(* IEC 61131-3 sources: 2026_Projet_YGO_ExcavatriceDragage/CODE/ENCODERS, 5 files *)

(* ---- ST_EncoderCalib.st ---- *)
(* ═══════════════════════════════════════════════════════════════
   🧲 ST_EncoderCalib — Calibration/référence codeur (1 par treuil, RETAIN)
   ───────────────────────────────────────────────────────────────
   📄 Doc métier : DOC/AF_Partie10_Fonction_Encoder_Homing_v1.6.md §9
   🎛️ Une instance RETAIN par treuil (M1_EncoderCalib / M2_EncoderCalib).
   ⚠️ Ce lot (acquisition + mise à l'échelle) : `HomingRefRaw` reste
      modifiable MANUELLEMENT (RETAIN, valeur de test) tant que
      `FB_Encoder_Homing` (qui l'écrit normalement, §5) n'est pas codé —
      même principe que le stub GVL du lot Winch.
   ═══════════════════════════════════════════════════════════════ *)

TYPE ST_EncoderCalib :
STRUCT
    HomingRefRaw                  : UDINT;   // Valeur brute figée au dernier homing réussi
    LastKnownRawPos                : UDINT;   // Dernier point brut valide connu (§3.7, continu)
    RestartCoherenceTolerancePts    : UDINT := 1000;  // Tolérance redémarrage (~12% PointsPerRev 8192)
    Homed                          : BOOL;    // TRUE dès qu'un référencement a réussi
    HomingSuspect                  : BOOL;    // TRUE si incohérence détectée au redémarrage (§3.7)
END_STRUCT
END_TYPE

(* ---- FB_Encoder_Abs.st ---- *)
(* ═══════════════════════════════════════════════════════════════
   🧲 FB_Encoder_Abs — Acquisition codeur absolu (accès bus, 1 responsabilité)
   ───────────────────────────────────────────────────────────────
   📄 Doc métier : DOC/AF_Partie10_Fonction_Encoder_Homing_v1.6.md §3/§6
   ⚠️ RÉÉCRITURE COMPLÈTE (remplace la version legacy du projet, dossier
      CODEUR) : l'ancienne version utilisait `HomingTrigger` (recalage
      instantané par simple offset) + un mode `Teach` auto-calibré —
      **incompatibles** avec le design Partie10 (preset SDO avec
      accusé, formule `CableM_PerRev` fixe). Retirés : `HomingTrigger`,
      `WaterLevelOffset`, `TeachActive/StartRaw/EndRaw/RealDistance`.
   🧩 1 FB = 1 responsabilité : accès bus EtherCAT + séquence d'écriture
      preset. N'orchestre PAS le homing lui-même (ça sera le rôle de
      `FB_Encoder_Homing`, pas codé ce lot) — `PresetRequest`/`PresetValue`
      sont pilotés en dur (`FALSE`/`0`) dans `PRG_MAIN` pour l'instant.
   🧊 Principe « geler sur doute » (§6) : `RawPos`/`AngleRaw`/`TurnCount`
      ne sont PAS mis à jour si `EncoderAvailable = FALSE` — ils
      conservent leur dernière valeur plausible.
   ✅ SÉQUENCE PRESET (§5) — CONFIRMÉ TERRAIN 2026-07-02 : `PresetTriggerCmd := 2`
      (valeur de commande, pas un masque de bits) déclenche le
      référencement du codeur à `PresetValueOut`. `CodeSeqTriggerCmd`
      (canal réel `COD1_CodeSeqTrigCmd`) reste `0`, rôle **non identifié**
      (même par l'utilisateur/terrain) — ne jamais lui donner une valeur
      arbitraire tant que sa fonction n'est pas confirmée.
   🔴 PERTE DE FONCTION SIGNALÉE : l'ancienne version composait
      `FB_Encoder_Safety` en interne (survitesse via `In_SpdValue`).
      Ce n'est PAS repris ici (Partie10 ne le demande pas, hors
      périmètre du document) — `FB_Encoder_Safety` (overspeed) devient
      orphelin tant qu'un lot dédié ne décide pas de son sort (fusion
      avec le "saut incohérent" Partie10 §3.5, ou reprise telle quelle).
   🔧 CORRECTIF (2026-07-03, retour terrain) : `InvertDirection` **retiré**.
      Confirmé terrain : l'objet CoE `6000h` (bit0 : 4→5) inverse le sens
      de comptage **côté codeur** (F58x8 Kübler), configuré en **Startup
      Parameter** CODESYS (init automate) — pas un paramètre PLC. L'ancien
      calcul logiciel (`16#FFFFFFFF - RawPosIn`) était de toute façon
      **buggé** : il inversait sur toute la plage `UDINT` (32 bits) au
      lieu de la plage réelle du codeur (25 bits, `PointsPerRev ×
      MultiTurnRevsMax`), produisant des positions incohérentes après
      homing. Voir Partie10 §3bis.
   ═══════════════════════════════════════════════════════════════ *)

// === DECLARATION (à coller dans la partie déclaration du POU FB_Encoder_Abs) ===

FUNCTION_BLOCK PUBLIC FB_Encoder_Abs
VAR_INPUT
    Enable              : BOOL;        // Standard
    Reset               : BOOL;        // Acquittement défaut (front)
    EmergencyStopOk     : BOOL;        // Standard
    Mode                : E_Mode;      // Standard (contexte, pas encore exploité ce lot)
    RawPosIn            : UDINT;       // Brut EtherCAT (ex. COD1_PosValue, %ID)
    AlarmsIn            : UINT;        // Brut EtherCAT (ex. COD1_Alarms)
    WarningsIn          : UINT;        // Brut EtherCAT (ex. COD1_Warnings) — informatif seulement
    SlaveOperational    : BOOL;        // FB_DiagEthercat — esclave EtherCAT opérationnel
    PointsPerRev        : UDINT := 8192;  // Résolution codeur confirmée (Partie10 §3.3)
    PresetRequest       : BOOL;        // Front — piloté par FB_Encoder_Homing (stub FALSE ce lot)
    PresetValue         : UDINT;       // Cible brute — piloté par FB_Encoder_Homing (stub 0 ce lot)
    PresetTimeout       : TIME := T#2s;
    PresetTolerancePts  : UDINT := 10; // Tolérance relecture post-preset
END_VAR
VAR_OUTPUT
    Ready               : BOOL;
    Busy                : BOOL;
    Done                : BOOL;
    Error               : BOOL;
    ErrorId             : WORD;        // bit0: "Défaut communication codeur" - alarme/bus codeur ; bit1: "Erreur référencement (timeout)" - preset refusé/timeout
    State               : E_State;
    StateAtError        : E_State;
    RawPos              : UDINT;       // Position brute — GELÉE si EncoderAvailable=FALSE
    EncoderAvailable    : BOOL;
    AngleRaw            : UINT;        // Informatif maintenance : RawPos MOD PointsPerRev
    TurnCount           : UDINT;       // Informatif maintenance : RawPos / PointsPerRev
    PresetAck           : BOOL;        // Pulse 1 cycle — écriture confirmée
    PresetNak           : BOOL;        // Pulse 1 cycle — écriture refusée/timeout
    PresetTriggerCmd    : WORD;        // → à câbler sur COD_PresettTrigCmd (RxPDO)
    CodeSeqTriggerCmd   : WORD;        // → à câbler sur COD_CodeSeqTrigCmd (RxPDO)
    PresetValueOut      : UDINT;       // → à câbler sur COD_PresetValue (RxPDO)
END_VAR
VAR
    ResetEdge           : R_TRIG;
    ErrorEdge           : R_TRIG;
    PresetReqEdge       : R_TRIG;
    PresetTimer         : TON;
    PresetSeqStep       : INT;         // 0=IDLE, 1=pulse CodeSeq, 2=pulse Trig, 3=attente confirmation
    RawDiff             : DINT;
    PresetTimerVisual   : TON;         // Timer pour laisser le temps de voir l'impulsion (1.5s)
END_VAR

// === IMPLEMENTATION (à coller dans le corps ST du POU FB_Encoder_Abs) ===

// 🛑 1. GATE
IF NOT Enable THEN
    EncoderAvailable := FALSE;
    State := E_State.DISABLED;
    Ready := FALSE; Busy := FALSE; Done := FALSE;
    PresetTriggerCmd := 16#0000; CodeSeqTriggerCmd := 16#0000; PresetValueOut := 0;
    PresetSeqStep := 0;
    PresetTimer(IN := FALSE, PT := PresetTimeout);
    PresetTimerVisual(IN := FALSE, PT := T#500MS);
    RETURN;
END_IF;

Ready := TRUE;
State := E_State.READY;

// 🔑 2. RESET FRONT
ResetEdge(CLK := Reset);

// 🔍 3. DIAGNOSTIC BUS / ALARME
IF (AlarmsIn <> 0) OR NOT SlaveOperational THEN
    ErrorId := ErrorId OR 16#0001;
ELSIF ResetEdge.Q THEN
    ErrorId := ErrorId AND 16#FFFE;
END_IF;
EncoderAvailable := (ErrorId AND 16#0001) = 0;

// 📥 4. LECTURE POSITION — GELER SUR DOUTE (Partie10 §6)
// Si EncoderAvailable=FALSE : RawPos/AngleRaw/TurnCount conservent leur dernière valeur (pas de RETURN
// global ici pour ne pas geler aussi la séquence preset/l'état — seule la lecture est gelée).
IF EncoderAvailable THEN
    RawPos := RawPosIn;   // 🔧 2026-07-03 : sens de comptage géré côté codeur (CoE 6000h bit0,
                          // startup parameter CODESYS) — voir Partie10 §3bis. Plus de calcul ici.
    AngleRaw := UDINT_TO_UINT(RawPos MOD PointsPerRev);
    TurnCount := RawPos / PointsPerRev;
END_IF;

// 🔧 5. SÉQUENCE PRESET (écriture bus)
// ✅ Confirmé terrain (2026-07-02) : PresettTrigCmd := 2 déclenche le référencement à
//    PresetValue (valeur de commande, pas un masque de bits — corrige l'hypothèse initiale).
// 🔴 CodeSeqTrigCmd : rôle NON identifié (même par l'utilisateur/terrain) — laissé à 0,
//    PAS piloté tant que sa fonction n'est pas confirmée (fiche technique ou essai dédié).
//    Ne jamais lui donner une valeur arbitraire "au cas où".
PresetReqEdge(CLK := PresetRequest);
PresetAck := FALSE; PresetNak := FALSE; // pulses 1 cycle uniquement
CodeSeqTriggerCmd := 16#0000;           // 🔴 non piloté — rôle inconnu, voir note ci-dessus
CASE PresetSeqStep OF
    0: // IDLE
        PresetTriggerCmd := 0;
        IF PresetReqEdge.Q AND EncoderAvailable THEN
            PresetValueOut := PresetValue;
            PresetSeqStep := 1;
            PresetTimer(IN := TRUE, PT := PresetTimeout);
        END_IF;
    1: // Déclenchement preset (laissé actif pendant 0.5s pour confort visuel en simulation/bus)
        PresetTriggerCmd := 2;   // ✅ Valeur confirmée terrain — référence le codeur à PresetValueOut
        RawDiff := UDINT_TO_DINT(RawPos) - UDINT_TO_DINT(PresetValueOut);
        IF ABS(RawDiff) <= UDINT_TO_DINT(PresetTolerancePts) THEN
            PresetTimer(IN := FALSE, PT := PresetTimeout);
            PresetTimerVisual(IN := TRUE, PT := T#500MS);
            IF PresetTimerVisual.Q THEN
                PresetTriggerCmd := 0;
                PresetAck := TRUE;
                PresetSeqStep := 0;
                PresetTimerVisual(IN := FALSE, PT := T#500MS);
            END_IF;
        ELSIF PresetTimer.Q THEN
            PresetTriggerCmd := 0;
            PresetNak := TRUE;
            ErrorId := ErrorId OR 16#0002;
            PresetSeqStep := 0;
            PresetTimer(IN := FALSE, PT := PresetTimeout);
            PresetTimerVisual(IN := FALSE, PT := T#500MS);
        END_IF;
END_CASE;
IF ResetEdge.Q AND (PresetSeqStep = 0) THEN
    ErrorId := ErrorId AND 16#FFFD;
END_IF;

// 🧾 6. ERROR / STATEATERROR
Error := (ErrorId <> 16#0000);
ErrorEdge(CLK := Error);
IF ErrorEdge.Q THEN
    StateAtError := State;
END_IF;

Busy := (PresetSeqStep <> 0);
Done := PresetAck;

(* ---- FB_Encoder_Homing.st ---- *)
(* ═══════════════════════════════════════════════════════════════
   🎯 FB_Encoder_Homing — Référencement codeur, flux NOMINAL uniquement
   ───────────────────────────────────────────────────────────────
   📄 Doc métier : DOC/AF_Partie10_Fonction_Encoder_Homing_v1.6.md §1/§5/§7bis
   ⚠️ PÉRIMÈTRE DE CE LOT : flux **nominal** uniquement (capteur haut +
      bouton IHM, référencement à `TopSensorPositionM`, 1 instance par
      treuil, câblées sur le MÊME bouton IHM côté PRG_MAIN). Le flux
      **unitaire** (`WinchSelect`, cible libre `HomingTargetM`,
      `MAINT_N2`) n'est **pas** codé ici — dépend de `E_WinchSelect`/
      `FB_Modes`, pas encore construits.
   🔌 PAS un FB de mouvement (Partie3 §1bis) : il n'écrit qu'une valeur
      de calibration, le treuil étant déjà à l'arrêt confirmé. Pas de
      `StartStop`/`SafeStop`.
   🧮 Calcul (généralise le cas historique cible=0.00, Partie10 §3.2/§3.3) :
      - `PresetValue` = `HomingRefTargetNominal` = (PointsPerRev × MultiTurnRevsMax) / 2
        (constante, TOUJOURS la même — centre exact de la plage, marge anti-débordement)
      - `HomingRefRaw` = `PresetValue` − round(`TopSensorPositionM` × PointsPerRev / CableM_PerRev)
        (ainsi `CablePosM` = `TopSensorPositionM` exactement au moment du homing)
      ⚠️ ÉVOLUTION vs interface §5 d'origine : `HomingRefRaw` est ajouté en sortie explicite
      (le document original supposait implicitement `HomingRefRaw := PresetValue`, valable
      uniquement pour une cible à 0.00 — ne fonctionne plus avec une cible non nulle ≈12.50 m).
   🧊 `ST_EncoderCalib` géré en interne (`VAR RETAIN`) — expose `Homed`/`HomingSuspect`/
      `HomingRefRaw` en sortie pour les consommateurs (`FB_Encoder_Scale`).
   🔴 SIMPLIFICATIONS assumées pour ce lot (à documenter/lever plus tard si besoin) :
      - Les 2 instances (M1/M2) sont autonomes : le même bouton IHM pilote les deux `Home`
        simultanément (câblage PRG_MAIN), mais chacune valide/rejette SES PROPRES conditions
        indépendamment (pas d'attente mutuelle ni de synchro de déclenchement).
      - `ConfirmCoherence`/§3.7 (incohérence redémarrage) : implémenté a minima (bit9), mais
        non testé en conditions réelles de coupure secteur — à revalider.
   ═══════════════════════════════════════════════════════════════ *)

// === DECLARATION (à coller dans la partie déclaration du POU FB_Encoder_Homing) ===

FUNCTION_BLOCK PUBLIC FB_Encoder_Homing
VAR_INPUT
    Enable               : BOOL;        // Standard
    Reset                : BOOL;        // Acquittement défaut (front) — bits 0/2/3/4/5 (voir §ErrorId)
    EmergencyStopOk      : BOOL;        // Standard
    Mode                 : E_Mode;      // MAINT_N1 requis pour le flux nominal
    Home                 : BOOL;        // Demande de référencement (front, bouton IHM UNIQUE)
    ConfirmCoherence     : BOOL;        // Front — lève le doute §3.7 (bit9), sans réhoming complet
    TopPositionSensor    : BOOL;        // 🔧 2026-07-02 : capteur position haute UNIQUE, COMMUN aux 2 treuils
                                         // (les 2 câbles hissent ensemble le même ensemble mécanique) — câblé
                                         // IDENTIQUEMENT sur les instances M1 ET M2 (PAS un capteur par treuil),
                                         // voir PRG_MAIN.st
    TopSensorPositionM   : REAL := 8.5;   // Cible homing nominal (RETAIN site, voir Partie10 §7bis)
    FwdRevSpeedFeedbackOff : BOOL;      // 🔧 REX 2026-07-07 : retour unique "tous contacteurs sens+vitesse
                                         // retombés" CE TREUIL — arrêt confirmé (remplace ContactorFeedbackFwd/Rev)
    BrakeFeedback        : BOOL;        // Retour contacteur frein CE TREUIL (TRUE = relâché, FALSE = collé)
    RawPos               : UDINT;       // Sortie FB_Encoder_Abs (déjà gelée sur doute)
    EncoderAvailable     : BOOL;        // Sortie FB_Encoder_Abs
    PresetAck            : BOOL;        // Pulse — sortie FB_Encoder_Abs (écriture confirmée)
    PresetNak            : BOOL;        // Pulse — sortie FB_Encoder_Abs (écriture refusée/timeout)
    PointsPerRev         : UDINT := 8192;   // Confirmé fiche technique (Partie10 §3.3)
    MultiTurnRevsMax     : UDINT := 4096;   // Confirmé fiche technique (Partie10 §3.3)
    CableM_PerRev        : REAL := 2.0;     // Confirmé terrain 2026-07-02 (Partie10 §2)
END_VAR
VAR_OUTPUT
    Ready                : BOOL;
    Busy                 : BOOL;
    Done                 : BOOL;        // Pulse 1 cycle — référencement réussi (miroir PresetAck)
    Error                : BOOL;
    ErrorId              : WORD;        // Voir table de bits en en-tête de fichier / doc §5
    State                : E_State;
    StateAtError         : E_State;
    PresetRequest        : BOOL;        // Pulse → FB_Encoder_Abs.PresetRequest
    PresetValue          : UDINT;       // → FB_Encoder_Abs.PresetValue (= HomingRefTargetNominal)
    Homed                : BOOL;        // RETAIN interne, miroir Calib.Homed
    HomingSuspect        : BOOL;        // RETAIN interne, miroir Calib.HomingSuspect
    HomingRefRaw         : UDINT;       // RETAIN interne, miroir Calib.HomingRefRaw → FB_Encoder_Scale
END_VAR
VAR_IN_OUT
    Calib                : ST_EncoderCalib;   // Référence vers l'état persistant global (survit aux téléchargements)
END_VAR
VAR
    ResetEdge            : R_TRIG;
    ErrorEdge            : R_TRIG;
    HomeEdge             : R_TRIG;
    ConfirmCoherenceEdge : R_TRIG;
    InitDone             : BOOL;        // Contrôle cohérence §3.7 fait une fois par session Enable
    ArretConfirme        : BOOL;
    PresetValueCalc      : UDINT;       // = HomingRefTargetNominal (constant tant que PointsPerRev/MultiTurnRevsMax fixes)
    TargetPoints         : DINT;        // Écart signé TopSensorPositionM → points, figé pendant la séquence
    RawDiffRestart       : DINT;        // Écart |RawPos - LastKnownRawPos| au redémarrage (§3.7)
END_VAR

// === IMPLEMENTATION (à coller dans le corps ST du POU FB_Encoder_Homing) ===

// 🛑 1. GATE — neutralisation ; on continue toutefois d'exposer le dernier état RETAIN connu
// (FB_Encoder_Scale a besoin de HomingRefRaw même si ce FB est désactivé)
IF NOT Enable THEN
    PresetRequest := FALSE;
    PresetValue := 0;
    State := E_State.DISABLED;
    Ready := FALSE; Busy := FALSE; Done := FALSE;
    InitDone := FALSE;   // Force un nouveau contrôle §3.7 à la prochaine activation
    Homed := Calib.Homed;
    HomingSuspect := Calib.HomingSuspect;
    HomingRefRaw := Calib.HomingRefRaw;
    RETURN;
END_IF;

Ready := TRUE;

// 🔑 2. FRONTS
ResetEdge(CLK := Reset);
HomeEdge(CLK := Home);
ConfirmCoherenceEdge(CLK := ConfirmCoherence);

// 🔍 3. COHÉRENCE AU REDÉMARRAGE (§3.7) — une fois par session Enable, dès que le codeur répond
IF NOT InitDone THEN
    State := E_State.INIT;
    IF EncoderAvailable THEN
        RawDiffRestart := UDINT_TO_DINT(RawPos) - UDINT_TO_DINT(Calib.LastKnownRawPos);
        IF Calib.Homed AND (ABS(RawDiffRestart) > UDINT_TO_DINT(Calib.RestartCoherenceTolerancePts)) THEN
            Calib.HomingSuspect := TRUE;
            ErrorId := ErrorId OR 16#0200;   // bit9 : incohérence codeur au redémarrage
        END_IF;
        InitDone := TRUE;
    END_IF;
ELSE
    IF State = E_State.INIT THEN State := E_State.READY; END_IF;
END_IF;

// ✅ 4. LEVÉE DU DOUTE (ConfirmCoherence, §3.7) — indépendant du Reset générique
IF ConfirmCoherenceEdge.Q AND (Mode = E_Mode.MAINT_N1 OR Mode = E_Mode.MAINT_N2) THEN
    Calib.HomingSuspect := FALSE;
    ErrorId := ErrorId AND 16#FDFF;   // efface bit9
END_IF;

// 🎯 5. DEMANDE DE RÉFÉRENCEMENT (flux nominal)
// ⚠️ `TopSensorPositionM` n'est PAS revalidée contre le bornage [-99.00;+99.00] m (§3.6) dans ce
// lot : c'est un paramètre RETAIN de mise en service (comme CableM_PerRev/PointsPerRev), pas une
// saisie opérateur par requête — valeur indicative ≈12.50 m largement dans la plage.
// 🔧 REX 2026-07-07 : FwdRevSpeedFeedbackOff remplace (NOT ContactorFeedbackFwd) AND (NOT ContactorFeedbackRev)
ArretConfirme := FwdRevSpeedFeedbackOff AND BrakeFeedback;

PresetRequest := FALSE;   // Défaut chaque cycle — repose uniquement sur le front HomeEdge ci-dessous
IF HomeEdge.Q AND (State <> E_State.BUSY) THEN
    // ✅ Homing autorisé en MAINT_N1 et MAINT_N2 — interdit en SEMI_AUTO et en cycle AUTO
    IF (Mode <> E_Mode.MAINT_N1) AND (Mode <> E_Mode.MAINT_N2) THEN
        ErrorId := ErrorId OR 16#0001;        // bit0 : mode non autorisé (seulement MAINT N1/N2)
    ELSIF NOT EncoderAvailable THEN
        ErrorId := ErrorId OR 16#0008;        // bit3 : codeur indisponible
    ELSIF NOT ArretConfirme THEN
        ErrorId := ErrorId OR 16#0004;        // bit2 : arrêt non confirmé (contacteurs/frein)
    ELSIF (Mode <> E_Mode.MAINT_N2) AND TopPositionSensor THEN
        // 🔧 CORRIGÉ 2026-07-04 : polarité inversée (testait NOT TopPositionSensor). Convention
        // NAMING_CONVENTION.md : TRUE = sain/non atteint, FALSE = position haute confirmée
        // (contact ouvert) — le Home nominal doit être rejeté tant que TopPositionSensor=TRUE.
        ErrorId := ErrorId OR 16#0010;        // bit4 : capteur position haute non confirmé (requis uniquement en MAINT_N1)
    ELSE
        // ✅ Toutes conditions réunies : calcul de la cible brute et déclenchement
        PresetValueCalc := (PointsPerRev * MultiTurnRevsMax) / 2;               // Centre exact (§3.3)
        TargetPoints := REAL_TO_DINT(TopSensorPositionM * UDINT_TO_REAL(PointsPerRev) / CableM_PerRev);
        PresetValue := PresetValueCalc;
        PresetRequest := TRUE;                // Pulse 1 cycle — FB_Encoder_Abs détecte le front lui-même
        State := E_State.BUSY;
    END_IF;
END_IF;

// ⏳ 6. SUIVI DE LA SÉQUENCE (BUSY → confirmation)
Done := FALSE;
IF State = E_State.BUSY THEN
    IF PresetAck THEN
        Calib.HomingRefRaw := DINT_TO_UDINT(UDINT_TO_DINT(PresetValueCalc) - TargetPoints);
        Calib.Homed := TRUE;
        Calib.HomingSuspect := FALSE;
        Calib.LastKnownRawPos := PresetValueCalc;
        Done := TRUE;
        State := E_State.READY;
        // 🔧 REX 2026-07-07 : un homing réussi re-établit la référence tout aussi validement
        // qu'un ConfirmCoherence explicite — efface donc aussi bit9 (incohérence redémarrage),
        // sinon ErrorId/Error restait bloqué à TRUE après un homing réussi (jamais mappé vers
        // l'IHM, invisible sauf sur GVL_IHM.Modes.AnyFaultActive qui restait à 1 sans raison visible).
        ErrorId := ErrorId AND 16#FDFF;
    ELSIF PresetNak THEN
        ErrorId := ErrorId OR 16#0020;        // bit5 : preset refusé/timeout (voir FB_Encoder_Abs)
        State := E_State.READY;
    END_IF;
END_IF;

// 🧾 7. RESET (front) — efface les bits « dernière tentative rejetée » (pas de cause persistante
// à revérifier ici : le prochain Home réévalue toutes les conditions de zéro, voir §5)
IF ResetEdge.Q THEN
    ErrorId := ErrorId AND 16#FFC2;   // efface bits 0,2,3,4,5 (garde bit9, levé seulement par ConfirmCoherence/Home)
END_IF;

// 📤 8. SORTIES ÉTAT
Error := (ErrorId <> 16#0000);
ErrorEdge(CLK := Error);
IF ErrorEdge.Q THEN
    StateAtError := State;
END_IF;

// Mise à jour continue du point brut valide connu (hors séquence de homing elle-même)
IF EncoderAvailable AND (State <> E_State.BUSY) THEN
    Calib.LastKnownRawPos := RawPos;
END_IF;

Busy := (State = E_State.BUSY);
Homed := Calib.Homed AND NOT Calib.HomingSuspect; // 🆕 REX 2026-07-08 : Perd l'état homed si suspect (démarrage ou fonctionnement), restauré après ConfirmCoherence
HomingSuspect := Calib.HomingSuspect;
HomingRefRaw := Calib.HomingRefRaw;

(* ---- FB_Encoder_Safety.st ---- *)
(* ═══════════════════════════════════════════════════════════════
   🛡️ FB_Encoder_Safety — Bornage physique + relais incohérence redémarrage (1 par treuil)
   ───────────────────────────────────────────────────────────────
   📄 Doc métier : DOC/AF_Partie10_Fonction_Encoder_Homing_v1.6.md §3.6/§3.7
   🔌 FB STANDARD (Partie3 §1bis) : pas un FB de mouvement, pas de StartStop/SafeStop.
   🎯 PÉRIMÈTRE CE LOT (répond à l'incident CablePosM≈4096m après reset RETAIN) :
      - §3.6 Bornage absolu [-99.00 ; +99.00] m : `CablePosM` hors plage → valeur
        jugée IMPOSSIBLE, sortie `CablePosMSafe` GELÉE sur dernière valeur plausible
        (principe « geler sur doute », §6), ErrorId bit0.
      - §3.7 Relais de `HomingSuspect` (déjà détecté par `FB_Encoder_Homing`, jamais
        consommé nulle part avant ce lot) : ErrorId bit1.
      - `EncoderIncoherent` (= Error) → consommé par `FB_Modes` pour REFUSER
        `SEMI_AUTO` (reste possible de travailler en MAINT_N1/N2 pour re-référencer,
        voir échange utilisateur — PAS de SafeStop ici, ne bloque jamais le mouvement).
   🔴 HORS PÉRIMÈTRE CE LOT (Partie10 §3.5, reporté) : détection de saut EN COURS
      D'EXPLOITATION (plausibilité vitesse codeur, calcul sur cycles EtherCAT 4ms) —
      lot dédié à part entière, pas fait ici.
   ═══════════════════════════════════════════════════════════════ *)

// === DECLARATION (à coller dans la partie déclaration du POU FB_Encoder_Safety) ===

FUNCTION_BLOCK PUBLIC FB_Encoder_Safety
VAR_INPUT
    Enable           : BOOL;        // Standard
    Reset            : BOOL;        // Acquittement défaut (front) — bit0 uniquement (bit1 suit HomingSuspect, voir §7bis)
    EmergencyStopOk  : BOOL;        // Standard
    Mode             : E_Mode;      // Standard (contexte, pas encore exploité ce lot)
    CablePosM        : REAL;        // Sortie FB_Encoder_Scale DE CE TREUIL
    HomingSuspect    : BOOL;        // Sortie FB_Encoder_Homing DE CE TREUIL (§3.7, déjà calculé)
    PositionMinM     : REAL := -99.0;  // Bornage physique dur (Partie10 §3.6)
    PositionMaxM     : REAL := 99.0;
END_VAR
VAR_OUTPUT
    Ready            : BOOL;
    Busy             : BOOL;
    Done             : BOOL;
    Error            : BOOL;
    ErrorId          : WORD;        // bit0: "Position câble hors plage" - position hors plage physique ; bit1: "Incohérence position boot" - incohérence redémarrage (miroir HomingSuspect)
    State            : E_State;
    StateAtError     : E_State;
    CablePosMSafe    : REAL;        // CablePosM gelée sur dernière valeur plausible si hors plage
    EncoderIncoherent: BOOL;        // = Error — consommé par FB_Modes (refuse SEMI_AUTO)
END_VAR
VAR
    ResetEdge             : R_TRIG;
    ErrorEdge             : R_TRIG;
    LastPlausibleCablePosM: REAL;
END_VAR

// === IMPLEMENTATION (à coller dans le corps ST du POU FB_Encoder_Safety) ===

// 🛑 1. GATE — expose la dernière valeur plausible connue même désactivé
IF NOT Enable THEN
    Ready := FALSE; Busy := FALSE; Done := FALSE;
    State := E_State.DISABLED;
    CablePosMSafe := LastPlausibleCablePosM;
    EncoderIncoherent := FALSE;
    RETURN;
END_IF;

Ready := TRUE;
State := E_State.READY;

// 🔑 2. RESET FRONT
ResetEdge(CLK := Reset);

// 🔍 3. BORNAGE PHYSIQUE ABSOLU (§3.6) — bit0
IF (CablePosM < PositionMinM) OR (CablePosM > PositionMaxM) THEN
    ErrorId := ErrorId OR 16#0001;
ELSIF ResetEdge.Q THEN
    ErrorId := ErrorId AND 16#FFFE;
END_IF;

// 🔍 4. RELAIS INCOHÉRENCE REDÉMARRAGE (§3.7, calculée par FB_Encoder_Homing) — bit1
// Pas d'acquittement ici : la levée se fait via ConfirmCoherence/nouveau Home côté
// FB_Encoder_Homing (source), ce FB ne fait QUE relayer l'information pour FB_Modes.
IF HomingSuspect THEN
    ErrorId := ErrorId OR 16#0002;
ELSE
    ErrorId := ErrorId AND 16#FFFD;
END_IF;

// 🧊 5. GELER SUR DOUTE (§6) — CablePosMSafe ne suit PAS CablePosM si hors plage
IF (ErrorId AND 16#0001) = 16#0000 THEN
    LastPlausibleCablePosM := CablePosM;
END_IF;
CablePosMSafe := LastPlausibleCablePosM;

// 📤 6. SORTIES ÉTAT
Error := (ErrorId <> 16#0000);
ErrorEdge(CLK := Error);
IF ErrorEdge.Q THEN
    StateAtError := State;
END_IF;

EncoderIncoherent := Error;
Busy := FALSE;
Done := FALSE;

(* ---- FB_Encoder_Scale.st ---- *)
(* ═══════════════════════════════════════════════════════════════
   📏 FB_Encoder_Scale — Mise à l'échelle points → mètres (1 par treuil)
   ───────────────────────────────────────────────────────────────
   📄 Doc métier : DOC/AF_Partie10_Fonction_Encoder_Homing_v1.6.md §2/§3.1
   ⚠️ RÉÉCRITURE (remplace la version legacy) : formule FIXE
      `CablePosM = (RawPos − HomingRefRaw) × (CableM_PerRev/PointsPerRev)`
      — retire le mode `Teach` auto-calibré (`EnableTeach`/`StartTeachPos`/
      `EndTeachPos`/`RealDistMeters`) : `CableM_PerRev` est un paramètre
      RETAIN fixe (site), pas recalculé dynamiquement (Partie10 §2).
   🧮 Arithmétique signée sûre (§3.1) : conversion en DINT AVANT la
      soustraction (jamais soustraire deux UDINT directement — un
      résultat négatif reboucle silencieusement vers ~2³²).
   🧩 Brique de calcul pure — pas de gel/bornage ici : `RawPos` en
      entrée est déjà gelé par `FB_Encoder_Abs` (§6) ; le bornage
      physique absolu [-99;+99] m est la responsabilité de
      `FB_Encoder_Safety` (§3.6, pas dans ce lot), pas de celle-ci.
   ═══════════════════════════════════════════════════════════════ *)

// === DECLARATION (à coller dans la partie déclaration du POU FB_Encoder_Scale) ===

FUNCTION_BLOCK PUBLIC FB_Encoder_Scale
VAR_INPUT
    RawPos          : UDINT;       // Position brute (sortie FB_Encoder_Abs, déjà gelée sur doute)
    HomingRefRaw    : UDINT;       // Référence brute figée au dernier homing (ST_EncoderCalib)
    CableM_PerRev   : REAL := 2.0; // Câble déroulé par tour (périmètre tambour confirmé 2026-07-02, réglable site)
    PointsPerRev    : UDINT := 8192; // Résolution codeur confirmée (Partie10 §3.3)
END_VAR
VAR_OUTPUT
    CablePosM       : REAL;        // Position câble en mètres, signée (+ enroulé, − sous l'eau)
END_VAR
VAR
    RawDiff         : DINT;        // Écart signé RawPos - HomingRefRaw (§3.1)
END_VAR

// === IMPLEMENTATION (à coller dans le corps ST du POU FB_Encoder_Scale) ===

// 🧮 Écart signé sûr : conversion DINT AVANT soustraction (§3.1) — jamais l'inverse
RawDiff := UDINT_TO_DINT(RawPos) - UDINT_TO_DINT(HomingRefRaw);

// 📏 Formule fixe points → mètres (Partie10 §2)
IF PointsPerRev > 0 THEN
    CablePosM := DINT_TO_REAL(RawDiff) * (CableM_PerRev / UDINT_TO_REAL(PointsPerRev));
ELSE
    CablePosM := 0.0;   // Garde division par zéro (PointsPerRev mal configuré)
END_IF;
